(* IEC 61131-3 sources: STAR-PLC-Agent/results/raw/four_group_20261114/star_terra/SELF001/formal/attempt_0001, 1 file *)

(* ---- candidate.st ---- *)
FUNCTION_BLOCK FB_Task
VAR_INPUT
    Start : BOOL;
    Stop : BOOL;
    GuardClosed : BOOL;
END_VAR
VAR_OUTPUT
    Run : BOOL := FALSE;
END_VAR
VAR
    running : BOOL := FALSE;
END_VAR

IF Stop OR NOT GuardClosed THEN
    running := FALSE;
ELSIF Start THEN
    running := TRUE;
END_IF;

Run := running;
END_FUNCTION_BLOCK
